{attribute 'TcGenerated'}
{attribute 'no-analysis'}
{attribute 'linkalways'}
// This function has been automatically generated from the project information.
VAR_GLOBAL CONSTANT
	{attribute 'const_non_replaced'}
	stLibVersion_ATI_KOSTAL_AF2024_AUDI2026_TcProjectBase : ST_LibVersion := (iMajor := 1, iMinor := 1, iBuild := 0, iRevision := 2, nFlags := 0, sVersion := '1.1.0.2');
END_VAR

(* stored: Version 1.1.0.1, ProductVersion 3.1.4024.12
   GVL Global_Version: Id {f129f3b9-6401-4ebb-91ee-6759c026fb8f} *)
